FUNCTION_BLOCK LightControll (* Composite Function Block Type *)
  (* Standard: 61499-2 *)
  (* Version 0.0, 10/20/2026, macie, Schneider Electric, template *)
  PACKAGE Main;
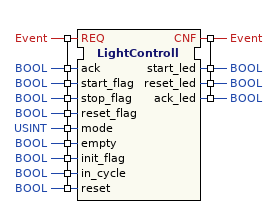
  EVENT_INPUT
    REQ WITH ack, start_flag, stop_flag, reset_flag, mode, empty, init_flag, in_cycle, reset; (* Normal Execution Request *)
  END_EVENT
  EVENT_OUTPUT
    CNF WITH start_led, reset_led, ack_led; (* Execution Confirmation *)
  END_EVENT
  VAR_INPUT
    ack : BOOL;
    start_flag : BOOL;
    stop_flag : BOOL;
    reset_flag : BOOL;
    mode : USINT;
    empty : BOOL;
    init_flag : BOOL;
    in_cycle : BOOL;
    reset : BOOL;
  END_VAR
  VAR_OUTPUT
    start_led : BOOL; (* Output event qualifier *)
    reset_led : BOOL;
    ack_led : BOOL;
  END_VAR
  FBS
    FB1 : StartLedControl;
    FB2 : ResetLedControl;
    FB3 : E_MERGE;
    FB4 : AckLedControl;
    FB5 : E_MERGE;
  END_FBS
  EVENT_CONNECTIONS
    REQ TO FB1.REQ;
    REQ TO FB2.REQ;
    FB1.CNF TO FB3.EI1;
    FB2.CNF TO FB3.EI2;
    FB3.EO TO FB5.EI1;
    FB4.CNF TO FB5.EI2;
    FB5.EO TO CNF;
    REQ TO FB4.REQ;
  END_CONNECTIONS
  DATA_CONNECTIONS
    stop_flag TO FB1.stop_flag;
    mode TO FB1.mode;
    start_flag TO FB1.start_flag;
    FB1.StartLed TO start_led;
    reset_flag TO FB1.reset_flag;
    empty TO FB1.empty;
    init_flag TO FB1.init_state;
    in_cycle TO FB1.in_cycle;
    stop_flag TO FB2.stop_flag;
    reset_flag TO FB2.reset_flag;
    mode TO FB2.mode;
    FB2.ResetLed TO reset_led;
    in_cycle TO FB2.in_cycle;
    start_flag TO FB2.start_flag;
    FB4.AckLed TO ack_led;
    empty TO FB4.empty;
    reset TO FB4.reset;
    ack TO FB4.ack;
  END_CONNECTIONS
END_FUNCTION_BLOCK
